SUBAPPLICATION Uebung_OPC_L12_AX (* Wie Training_12, lokal: Transport gebuendelt (A2X2_PUBLISH_2_SUBSCRIBE_2 statt CLIENT_2_0) *)
  (* Standard: 61499-2; Description: Copyright (c) 2026 Meisterschulen am Ostbahnhof This program and the accompanying materials are made available under the terms of the Eclipse Public License 2.0 which is available at https://www.eclipse.org/legal/epl-2.0/ SPDX-License-Identifier: EPL-2.0 *)
  (* Version 1.0, 2026-10-18, Franz Höpfinger, Meisterschulen am Ostbahnhof, Aus SubApp_PC_A + SubApp_PC_B von test_VV zusammengefuehrt, lokale Varianten der Bausteine *)
  PACKAGE Meins::OPC_UA_Lokal;
  IMPORT Uebungen::const::UT::DefaultPool::SoftKey_F1;
  IMPORT Uebungen::const::UT::DefaultPool::SoftKey_F2;
  IMPORT Meins::OPC_UA_Lokal::const::OpcUaLokal::SW2_PRESS_WRITE;
  IMPORT Meins::OPC_UA_Lokal::const::OpcUaLokal::SW2_STATE_READ;
  IMPORT Meins::OPC_UA_Lokal::const::OpcUaLokal::SW2_PRESS_READ;
  IMPORT Meins::OPC_UA_Lokal::const::OpcUaLokal::SW2_STATE_WRITE;
  IMPORT logiBUS::io::DQ::logiBUS_DO::Output_Q7;
  IMPORT logiBUS::io::DQ::logiBUS_DO::Output_Q8;
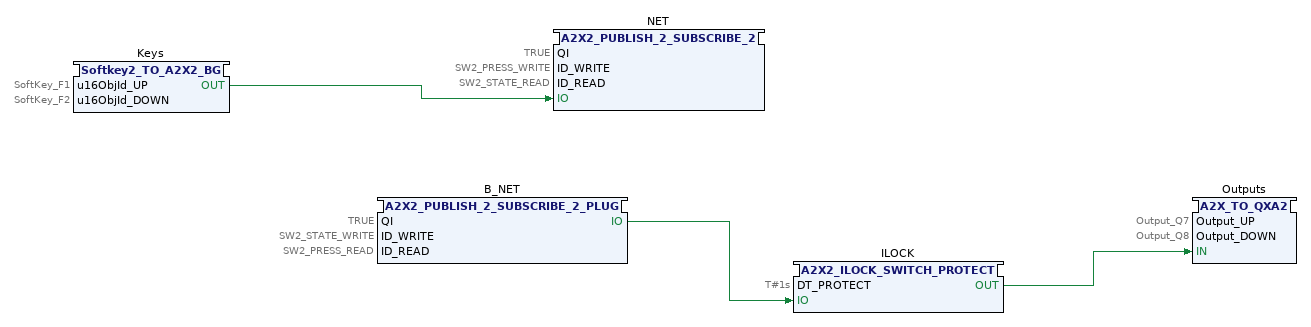
  SUBAPPS
    Keys : MyLib::sys::Softkey2_TO_A2X2_BG(u16ObjId_UP := SoftKey_F1, u16ObjId_DOWN := SoftKey_F2);
    NET : MyLib::net::A2X2_PUBLISH_2_SUBSCRIBE_2(QI := TRUE, ID_WRITE := SW2_PRESS_WRITE, ID_READ := SW2_STATE_READ);
    B_NET : MyLib::net::A2X2_PUBLISH_2_SUBSCRIBE_2_PLUG(QI := TRUE, ID_WRITE := SW2_STATE_WRITE, ID_READ := SW2_PRESS_READ);
    ILOCK : MyLib::sys::A2X2_ILOCK_SWITCH_PROTECT(DT_PROTECT := T#1s);
    Outputs : MyLib::sys::A2X_TO_QXA2(Output_UP := Output_Q7, Output_DOWN := Output_Q8);
  END_SUBAPPS
  ADAPTER_CONNECTIONS
    Keys.OUT TO NET.IO;
    B_NET.IO TO ILOCK.IO;
    ILOCK.OUT TO Outputs.IN;
  END_CONNECTIONS
END_SUBAPPLICATION
